(* Tests log record queue behavior and ownership transfer. *)
FUNCTION_BLOCK FB_TestLogRecordQueue EXTENDS FB_TestSuite

THIS^.testEnforcesMaximumSize();
THIS^.testAllowsUnboundedLength();
THIS^.testDropsOldestRecordFirst();
THIS^.testPushAndPopTransferRecordOwnership();
THIS^.testTransfersQueueOwnership();
THIS^.testTransfersRequestedCount();
THIS^.testReportsFailureReasons();

(* A queue built with maxCount 0 is unbounded and accepts every record without dropping; batch processors rely on this when no limit is configured. *)
METHOD testAllowsUnboundedLength : REFERENCE TO FB_Test
VAR
	queue: FB_LogRecordQueue(maxCount:=0);
	pRecord: POINTER TO FB_LogRecord;
	failureReason: E_LogRecordQueueFailureReason;
	success: BOOL;
	_idx: UDINT;
END_VAR
TcUnit.TEST('testAllowsUnboundedLength');
	FOR _idx := 1 TO 3 DO
		// opaque queue node: no factory hands a test an owned FB_LogRecord
		pRecord := __NEW(FB_LogRecord(severityNumber:=E_SeverityNumber.INFO, timestamp:=_idx));
		success := queue.push(pValue:=pRecord, failureReason=>failureReason);
		THIS^.AssertTrue(success AND_THEN pRecord = 0, 'Expected the unbounded queue to take ownership');
	END_FOR
	THIS^.AssertEquals_UDINT(3, queue.count, 'Expected maxSize zero to allow every record');
	THIS^.AssertEquals_UDINT(0, queue.droppedCount, 'Expected the unbounded queue not to drop records');
	queue.free();
TcUnit.TEST_FINISHED();
END_METHOD

(* A full queue drops its oldest record to make room for a new one, so the most recent logs survive a burst. *)
METHOD testDropsOldestRecordFirst : REFERENCE TO FB_Test
VAR
	queue: FB_LogRecordQueue(maxCount:=2);
	pRecord: POINTER TO FB_LogRecord;
	failureReason: E_LogRecordQueueFailureReason;
	success: BOOL;
	_idx: UDINT;
END_VAR
TcUnit.TEST('testDropsOldestRecordFirst');
	FOR _idx := 1 TO 3 DO
		// opaque queue node: no factory hands a test an owned FB_LogRecord
		pRecord := __NEW(FB_LogRecord(severityNumber:=E_SeverityNumber.INFO, timestamp:=_idx));
		success := queue.push(pValue:=pRecord, failureReason=>failureReason);
		THIS^.AssertTrue(success, 'Expected push to succeed');
	END_FOR

	success := queue.pop(pValue:=pRecord, failureReason=>failureReason);
	THIS^.AssertTrue(success AND_THEN pRecord <> 0 AND_THEN pRecord^.timestamp = 2, 'Expected timestamp 1 to be dropped first');
	IF pRecord <> 0 THEN pRecord^.delete(pSelf:=pRecord); END_IF
	success := queue.pop(pValue:=pRecord, failureReason=>failureReason);
	THIS^.AssertTrue(success AND_THEN pRecord <> 0 AND_THEN pRecord^.timestamp = 3, 'Expected the newest record to remain at the tail');
	IF pRecord <> 0 THEN pRecord^.delete(pSelf:=pRecord); END_IF
TcUnit.TEST_FINISHED();
END_METHOD

(* A bounded queue never holds more than maxCount records and counts each record it drops, so memory stays bounded on the PLC. *)
METHOD testEnforcesMaximumSize : REFERENCE TO FB_Test
VAR
	queue: FB_LogRecordQueue(maxCount:=2);
	pRecord: POINTER TO FB_LogRecord;
	failureReason: E_LogRecordQueueFailureReason;
	success: BOOL;
	_idx: UDINT;
END_VAR
TcUnit.TEST('testEnforcesMaximumSize');
	FOR _idx := 1 TO 3 DO
		// opaque queue node: no factory hands a test an owned FB_LogRecord
		pRecord := __NEW(FB_LogRecord(severityNumber:=E_SeverityNumber.INFO, timestamp:=_idx));
		success := queue.push(pValue:=pRecord, failureReason=>failureReason);
		THIS^.AssertTrue(success AND_THEN pRecord = 0, 'Expected push to take ownership');
		THIS^.AssertTrue(queue.count <= queue.maxCount, 'Expected count not to exceed maxSize');
	END_FOR
	THIS^.AssertTrue(queue.count = 2, 'Expected the queue to remain at its maximum size');
	THIS^.AssertTrue(queue.droppedCount = 1, 'Expected one record to be dropped');
TcUnit.TEST_FINISHED();
END_METHOD

(* Push takes ownership of the record and clears the caller's pointer, and pop hands the same record back; each record then has exactly one owner. *)
METHOD testPushAndPopTransferRecordOwnership : REFERENCE TO FB_Test
VAR
	queue: FB_LogRecordQueue(maxCount:=2);
	pRecord: POINTER TO FB_LogRecord;
	pOriginal: POINTER TO FB_LogRecord;
	failureReason: E_LogRecordQueueFailureReason;
	noFailure: E_LogRecordQueueFailureReason;
	success: BOOL;
END_VAR
TcUnit.TEST('testPushAndPopTransferRecordOwnership');
	noFailure := E_LogRecordQueueFailureReason.NA;
	// opaque queue node: no factory hands a test an owned FB_LogRecord
	pRecord := __NEW(FB_LogRecord(severityNumber:=E_SeverityNumber.INFO, timestamp:=42));
	pOriginal := pRecord;
	success := queue.push(pValue:=pRecord, failureReason=>failureReason);
	THIS^.AssertTrue(success AND_THEN failureReason = noFailure, 'Expected push to succeed without a failure reason');
	THIS^.AssertTrue(pRecord = 0 AND_THEN queue.count = 1, 'Expected push to transfer ownership into the queue');

	success := queue.pop(pValue:=pRecord, failureReason=>failureReason);
	THIS^.AssertTrue(success AND_THEN failureReason = noFailure, 'Expected pop to succeed without a failure reason');
	THIS^.AssertTrue(pRecord = pOriginal AND_THEN queue.count = 0, 'Expected pop to transfer the same record back to the caller');
	IF pRecord <> 0 THEN pRecord^.delete(pSelf:=pRecord); END_IF
TcUnit.TEST_FINISHED();
END_METHOD

(* Push and pop refuse a null record, an empty queue and an already assigned destination with a distinct reason each, and a later success clears the reason. *)
METHOD testReportsFailureReasons : REFERENCE TO FB_Test
VAR
	queue: FB_LogRecordQueue(maxCount:=1);
	pRecord: POINTER TO FB_LogRecord;
	pAssigned: POINTER TO FB_LogRecord;
	failureReason: E_LogRecordQueueFailureReason;
	noFailure: E_LogRecordQueueFailureReason;
	success: BOOL;
END_VAR
TcUnit.TEST('testReportsFailureReasons');
	noFailure := E_LogRecordQueueFailureReason.NA;
	success := queue.push(pValue:=pRecord, failureReason=>failureReason);
	THIS^.AssertFalse(success, 'Expected a null record push to fail');
	THIS^.AssertTrue(failureReason = E_LogRecordQueueFailureReason.RECORD_POINTER_NULL, 'Expected the null record failure reason');

	success := queue.pop(pValue:=pRecord, failureReason=>failureReason);
	THIS^.AssertFalse(success, 'Expected an empty pop to fail');
	THIS^.AssertTrue(failureReason = E_LogRecordQueueFailureReason.QUEUE_EMPTY, 'Expected the empty queue failure reason');

	// opaque queue node: no factory hands a test an owned FB_LogRecord
	pAssigned := __NEW(FB_LogRecord(severityNumber:=E_SeverityNumber.INFO, timestamp:=2));
	success := queue.pop(pValue:=pAssigned, failureReason=>failureReason);
	THIS^.AssertFalse(success, 'Expected pop into an assigned pointer to fail');
	THIS^.AssertTrue(failureReason = E_LogRecordQueueFailureReason.DESTINATION_ALREADY_ASSIGNED, 'Expected the assigned destination failure reason');
	IF pAssigned <> 0 THEN pAssigned^.delete(pSelf:=pAssigned); END_IF

	pRecord := __NEW(FB_LogRecord(severityNumber:=E_SeverityNumber.INFO, timestamp:=5));
	success := queue.push(pValue:=pRecord, failureReason=>failureReason);
	THIS^.AssertTrue(success AND_THEN failureReason = noFailure, 'Expected success to clear the previous failure reason');
TcUnit.TEST_FINISHED();
END_METHOD

(* transferTo moves records to another queue without copying them and keeps their FIFO order, so a batch can be handed on without new allocations. *)
METHOD testTransfersQueueOwnership : REFERENCE TO FB_Test
VAR
	source: FB_LogRecordQueue(maxCount:=2);
	destination: FB_LogRecordQueue(maxCount:=2);
	pRecord: POINTER TO FB_LogRecord;
	pFirstOriginal: POINTER TO FB_LogRecord;
	pSecondOriginal: POINTER TO FB_LogRecord;
	failureReason: E_LogRecordQueueFailureReason;
	noFailure: E_LogRecordQueueFailureReason;
	success: BOOL;
	_idx: UDINT;
END_VAR
TcUnit.TEST('testTransfersQueueOwnership');
	noFailure := E_LogRecordQueueFailureReason.NA;
	FOR _idx := 1 TO 2 DO
		// opaque queue node: no factory hands a test an owned FB_LogRecord
		pRecord := __NEW(FB_LogRecord(severityNumber:=E_SeverityNumber.INFO, timestamp:=_idx));
		IF _idx = 1 THEN
			pFirstOriginal := pRecord;
		ELSE
			pSecondOriginal := pRecord;
		END_IF
		success := source.push(pValue:=pRecord, failureReason=>failureReason);
		THIS^.AssertTrue(success, 'Expected source push to succeed');
	END_FOR

	success := source.transferTo(destination:=destination, count:=2, failureReason=>failureReason);
	THIS^.AssertTrue(success AND_THEN failureReason = noFailure, 'Expected queue ownership transfer to succeed');
	THIS^.AssertTrue(source.count = 0 AND_THEN destination.count = 2, 'Expected only the destination to own the records');

	success := destination.pop(pValue:=pRecord, failureReason=>failureReason);
	THIS^.AssertTrue(success AND_THEN pRecord = pFirstOriginal AND_THEN pRecord^.timestamp = 1, 'Expected transfer to preserve the first allocation and FIFO order');
	IF pRecord <> 0 THEN pRecord^.delete(pSelf:=pRecord); END_IF
	success := destination.pop(pValue:=pRecord, failureReason=>failureReason);
	THIS^.AssertTrue(success AND_THEN pRecord = pSecondOriginal AND_THEN pRecord^.timestamp = 2, 'Expected destination to own the same tail allocation');
	IF pRecord <> 0 THEN pRecord^.delete(pSelf:=pRecord); END_IF
TcUnit.TEST_FINISHED();
END_METHOD

(* transferTo moves only the requested number of oldest records and leaves the rest in the source, so a processor can export part of its queue. *)
METHOD testTransfersRequestedCount : REFERENCE TO FB_Test
VAR
	source: FB_LogRecordQueue(maxCount:=3);
	destination: FB_LogRecordQueue(maxCount:=0);
	pRecord: POINTER TO FB_LogRecord;
	failureReason: E_LogRecordQueueFailureReason;
	noFailure: E_LogRecordQueueFailureReason;
	success: BOOL;
	_idx: UDINT;
END_VAR
TcUnit.TEST('testTransfersRequestedCount');
	noFailure := E_LogRecordQueueFailureReason.NA;
	FOR _idx := 1 TO 3 DO
		// opaque queue node: no factory hands a test an owned FB_LogRecord
		pRecord := __NEW(FB_LogRecord(severityNumber:=E_SeverityNumber.INFO, timestamp:=_idx));
		success := source.push(pValue:=pRecord, failureReason=>failureReason);
		THIS^.AssertTrue(success, 'Expected source push to succeed');
	END_FOR

	success := source.transferTo(destination:=destination, count:=2, failureReason=>failureReason);
	THIS^.AssertTrue(success AND_THEN failureReason = noFailure, 'Expected a partial queue transfer to succeed');
	THIS^.AssertTrue(source.count = 1 AND_THEN destination.count = 2, 'Expected the destination to take only the requested count');

	success := destination.pop(pValue:=pRecord, failureReason=>failureReason);
	THIS^.AssertTrue(success AND_THEN pRecord <> 0 AND_THEN pRecord^.timestamp = 1, 'Expected the destination to receive the oldest record first');
	IF pRecord <> 0 THEN pRecord^.delete(pSelf:=pRecord); END_IF
	success := destination.pop(pValue:=pRecord, failureReason=>failureReason);
	THIS^.AssertTrue(success AND_THEN pRecord <> 0 AND_THEN pRecord^.timestamp = 2, 'Expected the destination to receive a FIFO slice');
	IF pRecord <> 0 THEN pRecord^.delete(pSelf:=pRecord); END_IF
	success := source.pop(pValue:=pRecord, failureReason=>failureReason);
	THIS^.AssertTrue(success AND_THEN pRecord <> 0 AND_THEN pRecord^.timestamp = 3, 'Expected the source to retain the untransferred tail');
	IF pRecord <> 0 THEN pRecord^.delete(pSelf:=pRecord); END_IF
TcUnit.TEST_FINISHED();
END_METHOD

END_FUNCTION_BLOCK

(* stored: Version 1.1.0.1
   POU FB_TestLogRecordQueue: Id {eae354c2-9892-456a-97c2-fbf651a21392}, SpecialFunc None
   Method testAllowsUnboundedLength: Id {019ff837-5af1-7c2a-a12a-b45f8f7d24d0}
   Method testDropsOldestRecordFirst: Id {cf630375-dba4-48d5-9684-440330c5de11}
   Method testEnforcesMaximumSize: Id {3d15347b-a733-498c-969f-bd92e68843e9}
   Method testPushAndPopTransferRecordOwnership: Id {a62a9c43-350f-4e05-b17a-4a95998386c2}
   Method testReportsFailureReasons: Id {09515266-8060-41de-97d3-7b1f99aac163}
   Method testTransfersQueueOwnership: Id {fb6226eb-9608-4e3d-8cfa-65afca222a12}
   Method testTransfersRequestedCount: Id {f5b79060-62be-451f-b340-4783541a9eaf} *)
